TYPE ST_SpindlePreheat_1 :
STRUCT
	dwOverride				:DWORD;			(* Override is percent of total speed of spindle. The range of override is from 0%  to 100 %  of rated speed.*)
	tDuration					:TIME;				(* Duration time for current phase *)
	dwSpeedRpm			:DWORD;			(* Current speed RPM - Read Only *)
	otstDuration				:OTSTRUCT;			(* Duration time in OTSTRUCT - Read Only*)
END_STRUCT
END_TYPE

(* stored: Version 1.1.0.1, ProductVersion 3.1.4024.15
   DUT ST_SpindlePreheat_1: Id {965789d8-f43e-4ec6-ada8-919bf74ee07e} *)
